Staubli VAL3: copyPoint31.pgx

public program copyPoint31(string x_sKey, num x_nTarget, num x_nSource)
  local num l_i
begin
  //2024.12.23 add 增加点位索引
  trajTemp:tTrajItem[x_sKey].pPointItem[x_nSource].pPointRx=tTrajBuffer[x_sKey].pPointItem[x_nTarget].pPointRx
  trajTemp:tTrajItem[x_sKey].pPointItem[x_nSource].pPointRx[1]=tTrajBuffer[x_sKey].pPointItem[x_nTarget].pPointRx[1]
  trajTemp:tTrajItem[x_sKey].pPointItem[x_nSource].jJointRx=tTrajBuffer[x_sKey].pPointItem[x_nTarget].jJointRx
  trajTemp:tTrajItem[x_sKey].pPointItem[x_nSource].sID=tTrajBuffer[x_sKey].pPointItem[x_nTarget].sID
  trajTemp:tTrajItem[x_sKey].pPointItem[x_nSource].bMarked=tTrajBuffer[x_sKey].pPointItem[x_nTarget].bMarked
  trajTemp:tTrajItem[x_sKey].pPointItem[x_nSource].pInter=tTrajBuffer[x_sKey].pPointItem[x_nTarget].pInter
  trajTemp:tTrajItem[x_sKey].pPointItem[x_nSource].pParaItem.mMdesc=tTrajBuffer[x_sKey].pPointItem[x_nTarget].pParaItem.mMdesc
  trajTemp:tTrajItem[x_sKey].pPointItem[x_nSource].pParaItem.nMoveType=tTrajBuffer[x_sKey].pPointItem[x_nTarget].pParaItem.nMoveType
  trajTemp:tTrajItem[x_sKey].pPointItem[x_nSource].pParaItem.nActionIndex=tTrajBuffer[x_sKey].pPointItem[x_nTarget].pParaItem.nActionIndex
  trajTemp:tTrajItem[x_sKey].pPointItem[x_nSource].pParaItem.nPercentage=tTrajBuffer[x_sKey].pPointItem[x_nTarget].pParaItem.nPercentage
  trajTemp:tTrajItem[x_sKey].pPointItem[x_nSource].pParaItem.nDelay=tTrajBuffer[x_sKey].pPointItem[x_nTarget].pParaItem.nDelay
  trajTemp:tTrajItem[x_sKey].pPointItem[x_nSource].pParaItem.nSigValue=tTrajBuffer[x_sKey].pPointItem[x_nTarget].pParaItem.nSigValue
  trajTemp:tTrajItem[x_sKey].pPointItem[x_nSource].pParaItem.bSafePoint=tTrajBuffer[x_sKey].pPointItem[x_nTarget].pParaItem.bSafePoint
  for l_i = 0 to 2
    trajTemp:tTrajItem[x_sKey].pPointItem[x_nSource].pParaItem.iIfItem.nSigType[l_i]=tTrajBuffer[x_sKey].pPointItem[x_nTarget].pParaItem.iIfItem.nSigType[l_i]
    trajTemp:tTrajItem[x_sKey].pPointItem[x_nSource].pParaItem.iIfItem.nSigIndex[l_i]=tTrajBuffer[x_sKey].pPointItem[x_nTarget].pParaItem.iIfItem.nSigIndex[l_i]
    trajTemp:tTrajItem[x_sKey].pPointItem[x_nSource].pParaItem.iIfItem.nValue[l_i]=tTrajBuffer[x_sKey].pPointItem[x_nTarget].pParaItem.iIfItem.nValue[l_i]
  endFor
  trajTemp:tTrajItem[x_sKey].pPointItem[x_nSource].pParaItem.iIfItem.bANDOR[0]=tTrajBuffer[x_sKey].pPointItem[x_nTarget].pParaItem.iIfItem.bANDOR[0]
  trajTemp:tTrajItem[x_sKey].pPointItem[x_nSource].pParaItem.iIfItem.bANDOR[1]=tTrajBuffer[x_sKey].pPointItem[x_nTarget].pParaItem.iIfItem.bANDOR[1]

end
